SUBAPPLICATION NetEv_Install_Filter (* NmGetCfInfo: install nur bei Active/NewAddress und nur einmal, sonst RSP *)
  (* Standard: 61499-2; Description: Copyright (c) 2026 Meisterschulen am Ostbahnhof This program and the accompanying materials are made available under the terms of the Eclipse Public License 2.0 which is available at https://www.eclipse.org/legal/epl-2.0/ SPDX-License-Identifier: EPL-2.0 *)
  (* Version 1.0, 2026-11-17, Franz Höpfinger, Meisterschulen am Ostbahnhof, initial implementation *)
  PACKAGE MyLib::sys;
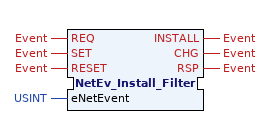
  EVENT_INPUT
    REQ; (* neues Netzwerkereignis *)
    SET; (* install erledigt (installO) *)
    RESET; (* wieder installieren erlauben *)
  END_EVENT
  EVENT_OUTPUT
    INSTALL; (* jetzt installieren *)
    CHG; (* schon installiert, Partner neu gemeldet (für CHG) *)
    RSP; (* nur quittieren (an NmGetCfInfo.RSP) *)
  END_EVENT
  VAR_INPUT
    eNetEvent : USINT; (* aus ISONETEVENT_T *)
  END_VAR
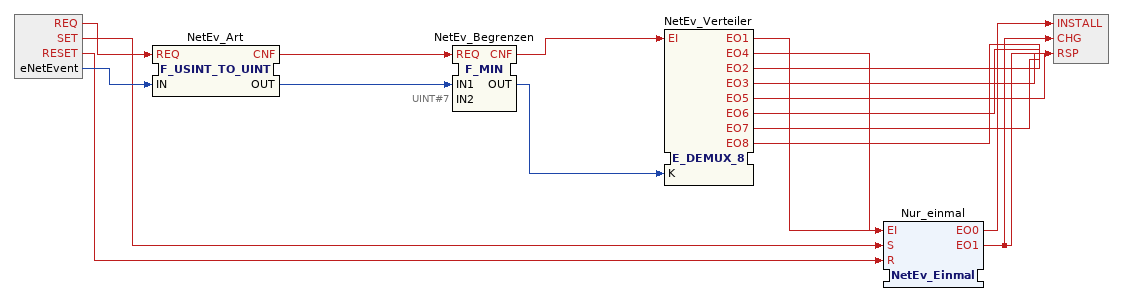
  FBS
    NetEv_Art : iec61131::conversion::F_USINT_TO_UINT;
    NetEv_Begrenzen : iec61131::selection::F_MIN(IN2 := UINT#7); (* ab 7 alles auf EO8, sonst kein RSP *)
    NetEv_Verteiler : iec61499::events::E_DEMUX_8(EO1 :=  (* Active *), EO2 :=  (* AddressConflict *), EO3 :=  (* Inactive *), EO4 :=  (* NewAddress *), EO5 :=  (* AddressViolation *), EO6 :=  (* MemberAdd *), EO7 :=  (* MemberRemove *), EO8 :=  (* 7 und mehr (Isonet_Last, HSI) *));
  END_FBS
  SUBAPPS
    Nur_einmal : MyLib::sys::NetEv_Einmal(EO0 :=  (* erstes Mal *), EO1 :=  (* schon erledigt *));
  END_SUBAPPS
  EVENT_CONNECTIONS
    REQ TO NetEv_Art.REQ;
    NetEv_Art.CNF TO NetEv_Begrenzen.REQ;
    NetEv_Begrenzen.CNF TO NetEv_Verteiler.EI;
    NetEv_Verteiler.EO1 TO Nur_einmal.EI;
    NetEv_Verteiler.EO4 TO Nur_einmal.EI;
    SET TO Nur_einmal.S;
    RESET TO Nur_einmal.R;
    Nur_einmal.EO0 TO INSTALL;
    Nur_einmal.EO1 TO CHG;
    Nur_einmal.EO1 TO RSP;
    NetEv_Verteiler.EO2 TO RSP;
    NetEv_Verteiler.EO3 TO RSP;
    NetEv_Verteiler.EO5 TO RSP;
    NetEv_Verteiler.EO6 TO RSP;
    NetEv_Verteiler.EO7 TO RSP;
    NetEv_Verteiler.EO8 TO RSP;
  END_CONNECTIONS
  DATA_CONNECTIONS
    eNetEvent TO NetEv_Art.IN;
    NetEv_Art.OUT TO NetEv_Begrenzen.IN1;
    NetEv_Begrenzen.OUT TO NetEv_Verteiler.K;
  END_CONNECTIONS
END_SUBAPPLICATION
